(* IEC 61131-3 sources: model-first-plc-agent-ai/results/T2-W-01, 2 files *)

(* ---- a1_code.st ---- *)
FUNCTION_BLOCK FB_TankFilling
VAR_INPUT
    start : BOOL;
    stop : BOOL;
    LSH : BOOL;
    LSHH : BOOL;
    TimerDuration : TIME;
END_VAR
VAR_OUTPUT
    fill_valve : BOOL;
    discharge_valve : BOOL;
END_VAR
VAR
    x0 : BOOL := TRUE;
    x1 : BOOL := FALSE;
    timer_done : BOOL := FALSE;
    fillingTimer : TON;
    t1_enabled : BOOL;
    t2_enabled : BOOL;
END_VAR

(* Evaluate elapsed time for the currently active filling step. *)
fillingTimer(IN := x1, PT := TimerDuration);
timer_done := fillingTimer.Q;

(* Evaluate both transitions against the same current situation. *)
t1_enabled := x0 AND start AND NOT stop AND NOT LSHH;
t2_enabled := x1 AND (stop OR LSHH OR timer_done);

IF t1_enabled THEN
    x0 := FALSE;
    x1 := TRUE;
ELSIF t2_enabled THEN
    x1 := FALSE;
    x0 := TRUE;
END_IF;

(* Start timing on entry and reset timing on exit in this scan. *)
IF t1_enabled OR t2_enabled THEN
    fillingTimer(IN := x1, PT := TimerDuration);
    timer_done := fillingTimer.Q;
END_IF;

fill_valve := x1;
discharge_valve := FALSE;

END_FUNCTION_BLOCK

PROGRAM Main
VAR
    StartCommand AT %IX100.0 : BOOL;
    StopCommand AT %IX100.1 : BOOL;
    LSH AT %IX100.2 : BOOL;
    LSHH AT %IX100.3 : BOOL;
    FillValve AT %QX100.0 : BOOL;
    DischargeValve AT %QX100.1 : BOOL;
END_VAR
VAR
    (* Configurable filling-time parameter; adjust for the scene. *)
    TimerDuration : TIME := T#10s;
    startEdge : R_TRIG;
    tankControl : FB_TankFilling;
END_VAR

startEdge(CLK := StartCommand);

tankControl(
    start := startEdge.Q,
    stop := StopCommand,
    LSH := LSH,
    LSHH := LSHH,
    TimerDuration := TimerDuration
);

FillValve := tankControl.fill_valve;
DischargeValve := tankControl.discharge_valve;

END_PROGRAM

(* ---- a2_code.st ---- *)
FUNCTION_BLOCK TankFillingController
VAR_INPUT
    StartCommand : BOOL;
    StopCommand : BOOL;
    LSH : BOOL;
    LSHH : BOOL;
    TimerDuration : TIME;
END_VAR
VAR_OUTPUT
    fill_valve : BOOL;
    discharge_valve : BOOL;
END_VAR
VAR
    ActiveStep : INT := 0;
    StartEdge : R_TRIG;
    FillingTimer : TON;
    start : BOOL;
    stop : BOOL;
    timer_done : BOOL;
END_VAR

StartEdge(CLK := StartCommand);
start := StartEdge.Q;
stop := StopCommand;

IF stop THEN
    ActiveStep := 0;
ELSE
    CASE ActiveStep OF
        0:
            IF start THEN
                ActiveStep := 1;
            END_IF;
        1:
            ActiveStep := 1;
    ELSE
        ActiveStep := 0;
    END_CASE;
END_IF;

(* Start timing in the same scan that the filling step becomes active. *)
FillingTimer(
    IN := (ActiveStep = 1),
    PT := TimerDuration
);
timer_done := FillingTimer.Q;

IF ActiveStep = 1 THEN
    IF stop OR timer_done OR LSHH THEN
        ActiveStep := 0;
    END_IF;
END_IF;

(* Reset the owned timer immediately upon leaving its step. *)
IF ActiveStep = 0 THEN
    FillingTimer(IN := FALSE, PT := TimerDuration);
    timer_done := FillingTimer.Q;
END_IF;

fill_valve := (ActiveStep = 1) AND NOT stop;
discharge_valve := FALSE;

END_FUNCTION_BLOCK

PROGRAM Main
VAR
    StartCommand AT %IX100.0 : BOOL;
    StopCommand AT %IX100.1 : BOOL;
    LSH AT %IX100.2 : BOOL;
    LSHH AT %IX100.3 : BOOL;
    FillValve AT %QX100.0 : BOOL;
    DischargeValve AT %QX100.1 : BOOL;
END_VAR
VAR
    Controller : TankFillingController;
    (* Configurable example preset; set to the required filling duration. *)
    TimerDuration : TIME := T#10s;
END_VAR

Controller(
    StartCommand := StartCommand,
    StopCommand := StopCommand,
    LSH := LSH,
    LSHH := LSHH,
    TimerDuration := TimerDuration
);

FillValve := Controller.fill_valve;
DischargeValve := Controller.discharge_valve;

END_PROGRAM
